(* IEC 61131-3 sources: ConveyorControl-with-PLC/4E_Gruppe1_Graf_Projekt1_HMI/Network, 1 file *)

(* ---- ConfigObjects.st ---- *)
FUNCTION GLOBAL TAB TASK_CONF
_K_TASK, _K_REAL,
_K_END_VAR,

_K_TASK, _K_CYCLIC,
_K_END_VAR,

_K_TASK, _K_BACKGROUND,
_K_END_VAR,

_K_END_CONF
END_FUNCTION

FUNCTION GLOBAL TAB IPR_CONF
_K_IPR
	0$UINT,
_K_END_VAR,
_K_END_CONF
END_FUNCTION

FUNCTION GLOBAL TAB CONFIG_TABLES
00030$UINT,
0$UINT, 0, 7, "_ALARMDISPLAY",
0$UINT, 0, 7, "_ALARMX0PARA",
0$UINT, 0, 2, "_ALARMX1PARA",
0$UINT, 0, 14, "_ALARMXBUFFER",
0$UINT, 0, 1, "_BIT32",
0$UINT, 0, 1, "_BIT32RAM",
0$UINT, 0, 12, "_GLOBAL",
0$UINT, 0, 1, "_HOTALARM",
0$UINT, 0, 4, "_LANGUAGESELECTION",
0$UINT, 0, 1, "_LIMITMAX",
0$UINT, 0, 1, "_LIMITMIN",
0$UINT, 0, 101, "_LSE",
0$UINT, 0, 3, "_MYIO",
0$UINT, 0, 6, "_OSZILSE",
0$UINT, 0, 0, "_OSZILSEBACKGROUND",
0$UINT, 0, 1, "_RADIO32",
0$UINT, 0, 1, "_RADIO32RAM",
0$UINT, 0, 2, "_SCREEN",
0$UINT, 0, 14, "_SCROLLAREA",
0$UINT, 0, 6, "_SCROLLAREA2",
0$UINT, 0, 5, "_SYSDATETIME",
0$UINT, 0, 2, "_TOOLCAT",
0$UINT, 0, 1, "_XACCESS",
0$UINT, 0, 10, "GETBROADCASTDATA",
0$UINT, 0, 1, "GRAPHIC",
0$UINT, 0, 6, "KEYPADANUM",
0$UINT, 0, 1, "KEYPADIMAGES",
0$UINT, 0, 3, "KEYPADNUM",
0$UINT, 1, 3, "RAM",
0$UINT, 0, 1, "SYSTEM",
ONE_CFG$UINT, 0, 0, "ONE_LseRtkAlarm",
ONE_CFG$UINT, 0, 0, "ONE_LseRtkMain",
TASK_CFG$UINT, 0, 0, "TASK_CONF",
IPR_CFG$UINT, 0, 0, "IPR_CONF",
PRJ_CFG$UINT, 0, 0, "4E_Gruppe1_Graf_Projekt1_HMI",
END_FUNCTION
